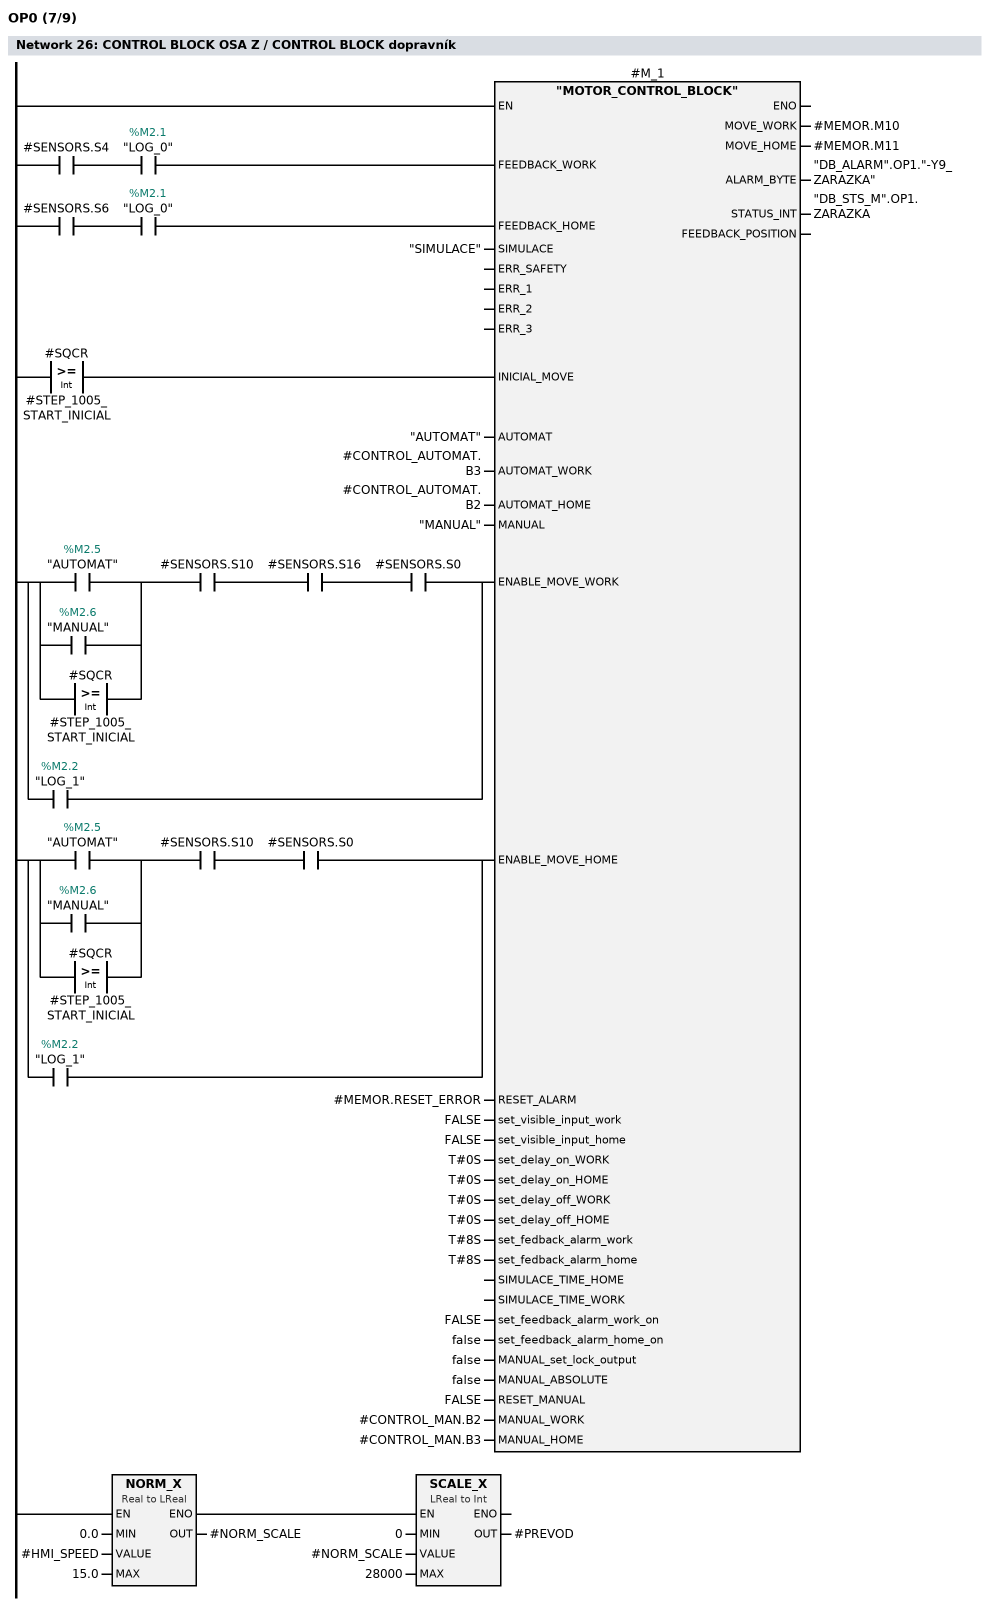
   RUNG wire#powerrail
      #M_1(FEEDBACK_WORK := wire#w1, FEEDBACK_HOME := wire#w2, INICIAL_MOVE := wire#w3, ENABLE_MOVE_WORK := wire#w5, ENABLE_MOVE_HOME := wire#w7, SIMULACE := "SIMULACE", ERR_SAFETY :=, ERR_1 :=, ERR_2 :=, ERR_3 :=, AUTOMAT := "AUTOMAT", AUTOMAT_WORK := #CONTROL_AUTOMAT.B3, AUTOMAT_HOME := #CONTROL_AUTOMAT.B2, MANUAL := "MANUAL", RESET_ALARM := #MEMOR.RESET_ERROR, set_visible_input_work := FALSE, set_visible_input_home := FALSE, set_delay_on_WORK := T#0S, set_delay_on_HOME := T#0S, set_delay_off_WORK := T#0S, set_delay_off_HOME := T#0S, set_fedback_alarm_work := T#8S, set_fedback_alarm_home := T#8S, SIMULACE_TIME_HOME :=, SIMULACE_TIME_WORK :=, set_feedback_alarm_work_on := FALSE, set_feedback_alarm_home_on := false, MANUAL_set_lock_output := false, MANUAL_ABSOLUTE := false, RESET_MANUAL := FALSE, MANUAL_WORK := #CONTROL_MAN.B2, MANUAL_HOME := #CONTROL_MAN.B3, MOVE_WORK => #MEMOR.M10, MOVE_HOME => #MEMOR.M11, ALARM_BYTE => "DB_ALARM".OP1."-Y9_ZARAZKA", STATUS_INT => "DB_STS_M".OP1.ZARAZKA, FEEDBACK_POSITION =>)
   END_RUNG
   RUNG wire#powerrail
      Contact( #SENSORS.S4 )
      Contact( "LOG_0" )
   END_RUNG wire#w1
   RUNG wire#powerrail
      Contact( #SENSORS.S6 )
      Contact( "LOG_0" )
   END_RUNG wire#w2
   RUNG wire#powerrail
      { S7_Templates := "SrcType := Int" } GE_Contact(in1 := #SQCR, in2 := #STEP_1005_START_INICIAL)
   END_RUNG wire#w3
   RUNG wire#powerrail
      Contact( "AUTOMAT" )
      wire#w4
      Contact( #SENSORS.S10 )
      Contact( #SENSORS.S16 )
      Contact( #SENSORS.S0 )
   END_RUNG wire#w5
   RUNG wire#powerrail
      Contact( "MANUAL" )
   END_RUNG wire#w4
   RUNG wire#powerrail
      { S7_Templates := "SrcType := Int" } GE_Contact(in1 := #SQCR, in2 := #STEP_1005_START_INICIAL)
   END_RUNG wire#w4
   RUNG wire#powerrail
      Contact( "LOG_1" )
   END_RUNG wire#w5
   RUNG wire#powerrail
      Contact( "AUTOMAT" )
      wire#w6
      Contact( #SENSORS.S10 )
      Contact( #SENSORS.S0 )
   END_RUNG wire#w7
   RUNG wire#powerrail
      Contact( "MANUAL" )
   END_RUNG wire#w6
   RUNG wire#powerrail
      { S7_Templates := "SrcType := Int" } GE_Contact(in1 := #SQCR, in2 := #STEP_1005_START_INICIAL)
   END_RUNG wire#w6
   RUNG wire#powerrail
      Contact( "LOG_1" )
   END_RUNG wire#w7
   RUNG wire#powerrail
      { S7_Templates := "[SrcType := Real, DestType := LReal]" } Normalize(min := 0.0, value := #HMI_SPEED, max := 15.0, out => #NORM_SCALE)
      { S7_Templates := "[SrcType := LReal, DestType := Int]" } Scale(min := 0, value := #NORM_SCALE, max := 28000, out => #PREVOD)
   END_RUNG
   // the same network as SCL:
   #M_1(FEEDBACK_WORK := #SENSORS.S4 AND "LOG_0",   // "MOTOR_CONTROL_BLOCK"
        FEEDBACK_HOME := #SENSORS.S6 AND "LOG_0",
        SIMULACE := "SIMULACE",
        INICIAL_MOVE := #SQCR >= #STEP_1005_START_INICIAL,
        AUTOMAT := "AUTOMAT",
        AUTOMAT_WORK := #CONTROL_AUTOMAT.B3,
        AUTOMAT_HOME := #CONTROL_AUTOMAT.B2,
        MANUAL := "MANUAL",
        ENABLE_MOVE_WORK := (("AUTOMAT" OR "MANUAL" OR (#SQCR >= #STEP_1005_START_INICIAL)) AND #SENSORS.S10 AND #SENSORS.S16 AND #SENSORS.S0) OR "LOG_1",
        ENABLE_MOVE_HOME := (("AUTOMAT" OR "MANUAL" OR (#SQCR >= #STEP_1005_START_INICIAL)) AND #SENSORS.S10 AND #SENSORS.S0) OR "LOG_1",
        RESET_ALARM := #MEMOR.RESET_ERROR,
        set_visible_input_work := FALSE,
        set_visible_input_home := FALSE,
        set_delay_on_WORK := T#0S,
        set_delay_on_HOME := T#0S,
        set_delay_off_WORK := T#0S,
        set_delay_off_HOME := T#0S,
        set_fedback_alarm_work := T#8S,
        set_fedback_alarm_home := T#8S,
        set_feedback_alarm_work_on := FALSE,
        set_feedback_alarm_home_on := false,
        MANUAL_set_lock_output := false,
        MANUAL_ABSOLUTE := false,
        RESET_MANUAL := FALSE,
        MANUAL_WORK := #CONTROL_MAN.B2,
        MANUAL_HOME := #CONTROL_MAN.B3,
        MOVE_WORK => #MEMOR.M10,
        MOVE_HOME => #MEMOR.M11,
        ALARM_BYTE => "DB_ALARM".OP1."-Y9_ZARAZKA",
        STATUS_INT => "DB_STS_M".OP1.ZARAZKA);
   #NORM_SCALE := NORM_X(MIN := 0.0, VALUE := #HMI_SPEED, MAX := 15.0);
   #PREVOD := SCALE_X(MIN := 0, VALUE := #NORM_SCALE, MAX := 28000);
END_REGION

REGION Network 27: CONTROL BLOCK ARETACE HLAVY / CONTROL BLOCK dveře laser
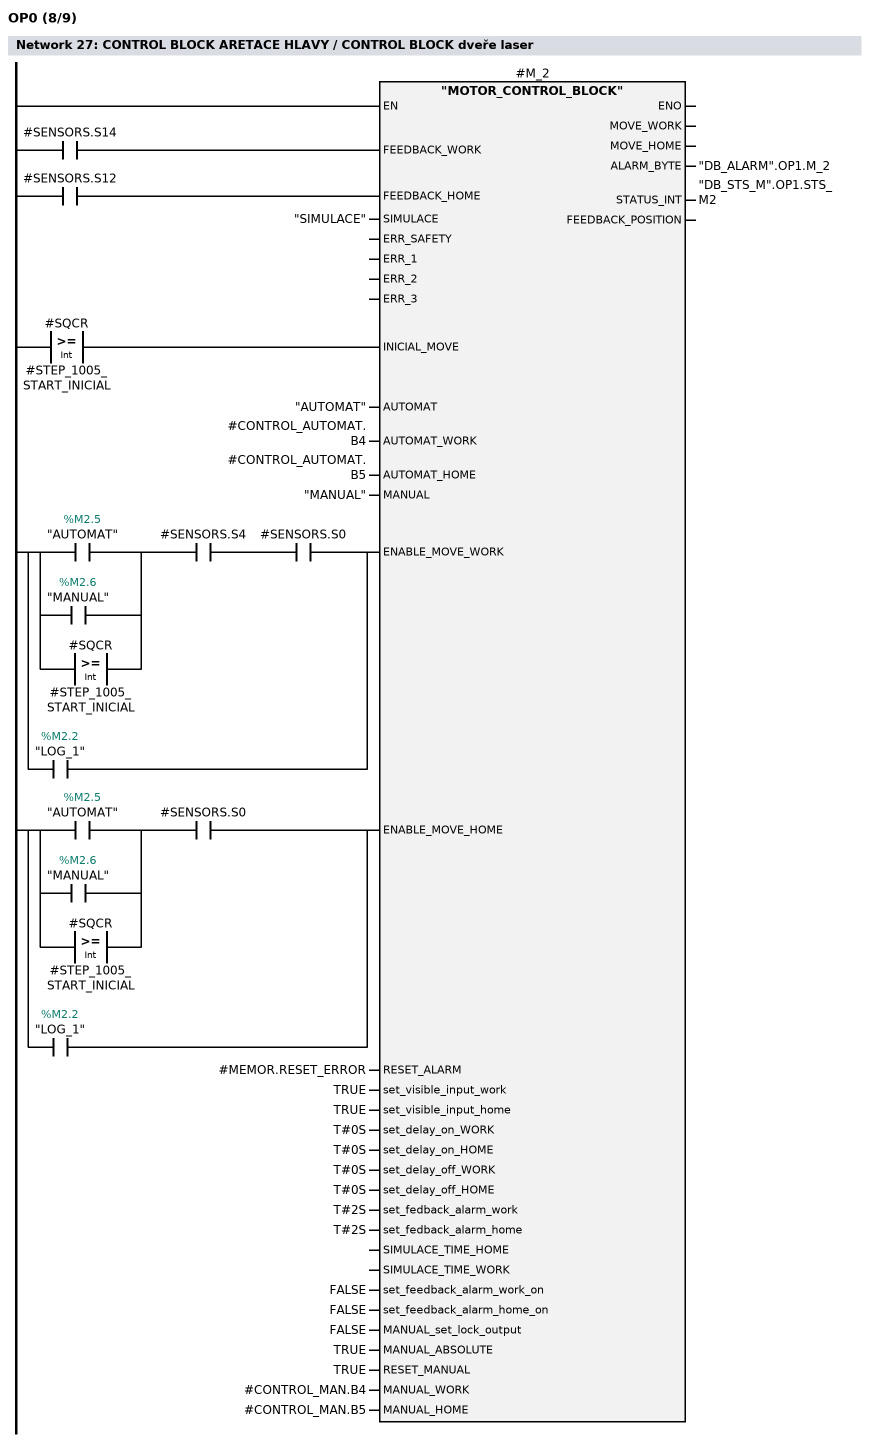
   RUNG wire#powerrail
      #M_2(FEEDBACK_WORK := wire#w1, FEEDBACK_HOME := wire#w2, INICIAL_MOVE := wire#w3, ENABLE_MOVE_WORK := wire#w5, ENABLE_MOVE_HOME := wire#w7, SIMULACE := "SIMULACE", ERR_SAFETY :=, ERR_1 :=, ERR_2 :=, ERR_3 :=, AUTOMAT := "AUTOMAT", AUTOMAT_WORK := #CONTROL_AUTOMAT.B4, AUTOMAT_HOME := #CONTROL_AUTOMAT.B5, MANUAL := "MANUAL", RESET_ALARM := #MEMOR.RESET_ERROR, set_visible_input_work := TRUE, set_visible_input_home := TRUE, set_delay_on_WORK := T#0S, set_delay_on_HOME := T#0S, set_delay_off_WORK := T#0S, set_delay_off_HOME := T#0S, set_fedback_alarm_work := T#2S, set_fedback_alarm_home := T#2S, SIMULACE_TIME_HOME :=, SIMULACE_TIME_WORK :=, set_feedback_alarm_work_on := FALSE, set_feedback_alarm_home_on := FALSE, MANUAL_set_lock_output := FALSE, MANUAL_ABSOLUTE := TRUE, RESET_MANUAL := TRUE, MANUAL_WORK := #CONTROL_MAN.B4, MANUAL_HOME := #CONTROL_MAN.B5, MOVE_WORK =>, MOVE_HOME =>, ALARM_BYTE => "DB_ALARM".OP1.M_2, STATUS_INT => "DB_STS_M".OP1.STS_M2, FEEDBACK_POSITION =>)
   END_RUNG
   RUNG wire#powerrail
      Contact( #SENSORS.S14 )
   END_RUNG wire#w1
   RUNG wire#powerrail
      Contact( #SENSORS.S12 )
   END_RUNG wire#w2
   RUNG wire#powerrail
      { S7_Templates := "SrcType := Int" } GE_Contact(in1 := #SQCR, in2 := #STEP_1005_START_INICIAL)
   END_RUNG wire#w3
   RUNG wire#powerrail
      Contact( "AUTOMAT" )
      wire#w4
      Contact( #SENSORS.S4 )
      Contact( #SENSORS.S0 )
   END_RUNG wire#w5
   RUNG wire#powerrail
      Contact( "MANUAL" )
   END_RUNG wire#w4
   RUNG wire#powerrail
      { S7_Templates := "SrcType := Int" } GE_Contact(in1 := #SQCR, in2 := #STEP_1005_START_INICIAL)
   END_RUNG wire#w4
   RUNG wire#powerrail
      Contact( "LOG_1" )
   END_RUNG wire#w5
   RUNG wire#powerrail
      Contact( "AUTOMAT" )
      wire#w6
      Contact( #SENSORS.S0 )
   END_RUNG wire#w7
   RUNG wire#powerrail
      Contact( "MANUAL" )
   END_RUNG wire#w6
   RUNG wire#powerrail
      { S7_Templates := "SrcType := Int" } GE_Contact(in1 := #SQCR, in2 := #STEP_1005_START_INICIAL)
   END_RUNG wire#w6
   RUNG wire#powerrail
      Contact( "LOG_1" )
   END_RUNG wire#w7
   // the same network as SCL:
   #M_2(FEEDBACK_WORK := #SENSORS.S14,   // "MOTOR_CONTROL_BLOCK"
        FEEDBACK_HOME := #SENSORS.S12,
        SIMULACE := "SIMULACE",
        INICIAL_MOVE := #SQCR >= #STEP_1005_START_INICIAL,
        AUTOMAT := "AUTOMAT",
        AUTOMAT_WORK := #CONTROL_AUTOMAT.B4,
        AUTOMAT_HOME := #CONTROL_AUTOMAT.B5,
        MANUAL := "MANUAL",
        ENABLE_MOVE_WORK := (("AUTOMAT" OR "MANUAL" OR (#SQCR >= #STEP_1005_START_INICIAL)) AND #SENSORS.S4 AND #SENSORS.S0) OR "LOG_1",
        ENABLE_MOVE_HOME := (("AUTOMAT" OR "MANUAL" OR (#SQCR >= #STEP_1005_START_INICIAL)) AND #SENSORS.S0) OR "LOG_1",
        RESET_ALARM := #MEMOR.RESET_ERROR,
        set_visible_input_work := TRUE,
        set_visible_input_home := TRUE,
        set_delay_on_WORK := T#0S,
        set_delay_on_HOME := T#0S,
        set_delay_off_WORK := T#0S,
        set_delay_off_HOME := T#0S,
        set_fedback_alarm_work := T#2S,
        set_fedback_alarm_home := T#2S,
        set_feedback_alarm_work_on := FALSE,
        set_feedback_alarm_home_on := FALSE,
        MANUAL_set_lock_output := FALSE,
        MANUAL_ABSOLUTE := TRUE,
        RESET_MANUAL := TRUE,
        MANUAL_WORK := #CONTROL_MAN.B4,
        MANUAL_HOME := #CONTROL_MAN.B5,
        ALARM_BYTE => "DB_ALARM".OP1.M_2,
        STATUS_INT => "DB_STS_M".OP1.STS_M2);
END_REGION

REGION Network 28: EXTERNAL_TRIGER
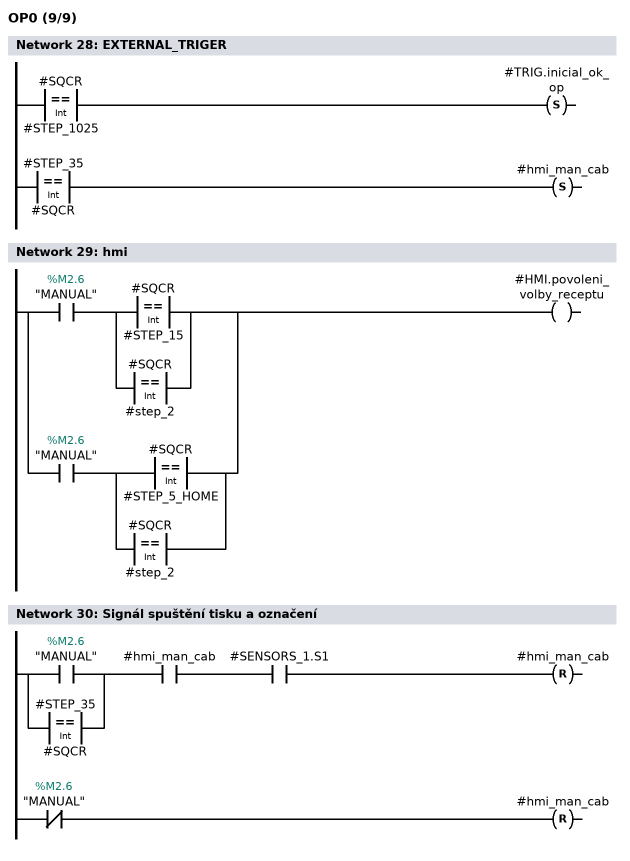
   RUNG wire#powerrail
      { S7_Templates := "SrcType := Int" } EQ_Contact(in1 := #SQCR, in2 := #STEP_1025)
      S_Coil( #TRIG.inicial_ok_op )
   END_RUNG
   RUNG wire#powerrail
      { S7_Templates := "SrcType := Int" } EQ_Contact(in1 := #STEP_35, in2 := #SQCR)
      S_Coil( #hmi_man_cab )
   END_RUNG
   // the same network as SCL:
   IF #SQCR = #STEP_1025 THEN #TRIG.inicial_ok_op := TRUE; END_IF;
   IF #STEP_35 = #SQCR THEN #hmi_man_cab := TRUE; END_IF;
END_REGION

REGION Network 29: hmi
   RUNG wire#powerrail
      Contact( "MANUAL" )
      wire#w1
      { S7_Templates := "SrcType := Int" } EQ_Contact(in1 := #SQCR, in2 := #STEP_15)
      wire#w2
      Coil( #HMI.povoleni_volby_receptu )
   END_RUNG
   RUNG wire#w1
      { S7_Templates := "SrcType := Int" } EQ_Contact(in1 := #SQCR, in2 := #step_2)
   END_RUNG wire#w2
   RUNG wire#powerrail
      Contact( "MANUAL" )
      wire#w3
      { S7_Templates := "SrcType := Int" } EQ_Contact(in1 := #SQCR, in2 := #STEP_5_HOME)
   END_RUNG wire#w2
   RUNG wire#w3
      { S7_Templates := "SrcType := Int" } EQ_Contact(in1 := #SQCR, in2 := #step_2)
   END_RUNG wire#w2
   // the same network as SCL:
   #HMI.povoleni_volby_receptu := ("MANUAL" AND ((#SQCR = #STEP_15) OR (#SQCR = #step_2))) OR ("MANUAL" AND ((#SQCR = #STEP_5_HOME) OR (#SQCR = #step_2)));
END_REGION

REGION Network 30: Signál spuštění tisku a označení
   RUNG wire#powerrail
      Contact( "MANUAL" )
      wire#w1
      Contact( #hmi_man_cab )
      Contact( #SENSORS_1.S1 )
      R_Coil( #hmi_man_cab )
   END_RUNG
   RUNG wire#powerrail
      { S7_Templates := "SrcType := Int" } EQ_Contact(in1 := #STEP_35, in2 := #SQCR)
   END_RUNG wire#w1
   RUNG wire#powerrail
      I_Contact( "MANUAL" )
      R_Coil( #hmi_man_cab )
   END_RUNG
   // the same network as SCL:
   IF ("MANUAL" OR (#STEP_35 = #SQCR)) AND #hmi_man_cab AND #SENSORS_1.S1 THEN #hmi_man_cab := FALSE; END_IF;
   IF NOT "MANUAL" THEN #hmi_man_cab := FALSE; END_IF;
END_REGION
END_FUNCTION_BLOCK

FUNCTION_BLOCK "OVLADANI_LASER"   // FB400, LAD
{ S7_Optimized_Access := 'TRUE' }
// stored: AutoNumber false, MemoryReserve 100, SetENOAutomatically false
   VAR
      SQCR : Int;
      SQCR_WHILE : Int;
      SET_WHILE : Bool;
      NAZEV_PROGRAMU : String[20];
      DELKA_STRINGU : Int;
      CHAR_K_ZAPISU : Array[0..71] of Char;
   END_VAR
   VAR CONSTANT
      STEP_0 : Int := 0;
      STEP_5 : Int := 5;
      STEP_10 : Int := 10;
      STEP_15 : Int := 15;
      STEP_20 : Int := 20;
      STEP_25 : Int := 25;
      STEP_30 : Int := 30;
      STEP_35 : Int := 35;
      STEP_40 : Int := 40;
      STEP_45 : Int := 45;
      STEP_50 : Int := 50;
      STEP_55 : Int := 55;
      STEP_60 : Int := 60;
      STEP_65 : Int := 65;
      STEP_70 : Int := 70;
      STEP_75 : Int := 75;
      STEP_80 : Int := 80;
      STEP_85 : Int := 85;
      STEP_90 : Int := 90;
      STEP_95 : Int := 95;
      STEP_100 : Int := 100;
   END_VAR
BEGIN

REGION Network 1
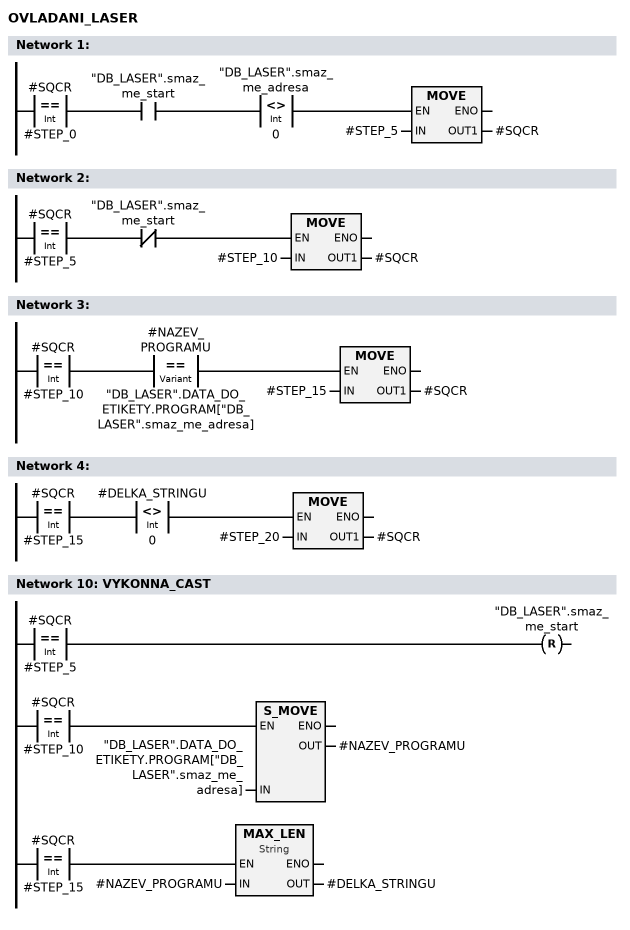
   RUNG wire#powerrail
      { S7_Templates := "SrcType := Int" } EQ_Contact(in1 := #SQCR, in2 := #STEP_0)
      Contact( "DB_LASER".smaz_me_start )
      { S7_Templates := "SrcType := Int" } NE_Contact(in1 := "DB_LASER".smaz_me_adresa, in2 := 0)
      Move(in := #STEP_5, out1 => #SQCR)
   END_RUNG
   // the same network as SCL:
   IF (#SQCR = #STEP_0) AND "DB_LASER".smaz_me_start AND ("DB_LASER".smaz_me_adresa <> 0) THEN
       #SQCR := #STEP_5;
   END_IF;
END_REGION

REGION Network 2
   RUNG wire#powerrail
      { S7_Templates := "SrcType := Int" } EQ_Contact(in1 := #SQCR, in2 := #STEP_5)
      I_Contact( "DB_LASER".smaz_me_start )
      Move(in := #STEP_10, out1 => #SQCR)
   END_RUNG
   // the same network as SCL:
   IF (#SQCR = #STEP_5) AND NOT "DB_LASER".smaz_me_start THEN #SQCR := #STEP_10; END_IF;
END_REGION

REGION Network 3
   RUNG wire#powerrail
      { S7_Templates := "SrcType := Int" } EQ_Contact(in1 := #SQCR, in2 := #STEP_10)
      { S7_Templates := "SrcType := Variant" } EQ_Contact(in1 := #NAZEV_PROGRAMU, in2 := "DB_LASER".DATA_DO_ETIKETY.PROGRAM["DB_LASER".smaz_me_adresa])
      Move(in := #STEP_15, out1 => #SQCR)
   END_RUNG
   // the same network as SCL:
   IF (#SQCR = #STEP_10) AND (#NAZEV_PROGRAMU = "DB_LASER".DATA_DO_ETIKETY.PROGRAM["DB_LASER".smaz_me_adresa]) THEN
       #SQCR := #STEP_15;
   END_IF;
END_REGION

REGION Network 4
   RUNG wire#powerrail
      { S7_Templates := "SrcType := Int" } EQ_Contact(in1 := #SQCR, in2 := #STEP_15)
      { S7_Templates := "SrcType := Int" } NE_Contact(in1 := #DELKA_STRINGU, in2 := 0)
      Move(in := #STEP_20, out1 => #SQCR)
   END_RUNG
   // the same network as SCL:
   IF (#SQCR = #STEP_15) AND (#DELKA_STRINGU <> 0) THEN #SQCR := #STEP_20; END_IF;
END_REGION

REGION Network 5: STEP_20 SCL NETVORK X
END_REGION

REGION Network 10: VYKONNA_CAST
   IF #SQCR = #STEP_5 THEN "DB_LASER".smaz_me_start := FALSE; END_IF;
   IF #SQCR = #STEP_10 THEN
       #NAZEV_PROGRAMU := "DB_LASER".DATA_DO_ETIKETY.PROGRAM["DB_LASER".smaz_me_adresa];
   END_IF;
   IF #SQCR = #STEP_15 THEN MAX_LEN(in := #NAZEV_PROGRAMU, out => #DELKA_STRINGU); END_IF;
END_REGION

REGION Network 12 (SCL)
   IF #SQCR = #STEP_20 THEN
       // zapsani počátečního znaku 
       #CHAR_K_ZAPISU[0] := "DB_LASER".DATA_DO_DAT.ZAVORKA_P;



       // vytvoření prdelky k názvu programu z laseru
       #CHAR_K_ZAPISU[#DELKA_STRINGU + 1] := "DB_LASER".DATA_DO_DAT.XLP[0];
       #CHAR_K_ZAPISU[#DELKA_STRINGU + 2] := "DB_LASER".DATA_DO_DAT.XLP[1];
       #CHAR_K_ZAPISU[#DELKA_STRINGU + 3] := "DB_LASER".DATA_DO_DAT.XLP[2];
       #CHAR_K_ZAPISU[#DELKA_STRINGU + 4] := "DB_LASER".DATA_DO_DAT.XLP[3];
       #CHAR_K_ZAPISU[#DELKA_STRINGU + 5] := "DB_LASER".DATA_DO_DAT.ZAVORKA_P;

       // dinamický zápis názvu podle délky stringu 
       WHILE #SET_WHILE DO
           IF #SQCR_WHILE > #DELKA_STRINGU THEN
               #SQCR_WHILE := 0;
               #SET_WHILE := FALSE;
               #SQCR := #STEP_25;
           ELSE
               #SQCR_WHILE := #SQCR_WHILE + 1;
           END_IF;
           #CHAR_K_ZAPISU[#SQCR_WHILE + 1] := #NAZEV_PROGRAMU[#SQCR_WHILE];
       END_WHILE;

   END_IF;
END_REGION
END_FUNCTION_BLOCK

FUNCTION "FC_PocetChyb" : Int
{ S7_Optimized_Access := 'TRUE' }
VERSION : 0.1
   VAR_INPUT 
      A : String;
      B : String;
   END_VAR

   VAR_TEMP 
      la : Int;
      lb : Int;
      i : Int;
      j : Int;
      v : Int;
      prev : Array[0..40] of Int;
      cur : Array[0..40] of Int;
   END_VAR


BEGIN
	// Pocet chyb mezi texty A a B (kolik znaku zamenit / vlozit / smazat).
	// 0 = texty jsou shodne. Porovnava se max. 40 znaku kvuli dobe cyklu.
	#la := MIN(IN1 := LEN(#A), IN2 := 40);
	#lb := MIN(IN1 := LEN(#B), IN2 := 40);
	
	FOR #j := 0 TO #lb DO
	    #prev[#j] := #j;
	END_FOR;
	
	FOR #i := 1 TO #la DO
	    #cur[0] := #i;
	    FOR #j := 1 TO #lb DO
	        #v := #prev[#j - 1];                // shoda / zamena znaku
	        IF #A[#i] <> #B[#j] THEN
	            #v := #v + 1;
	        END_IF;
	        IF #prev[#j] + 1 < #v THEN          // znak navic
	            #v := #prev[#j] + 1;
	        END_IF;
	        IF #cur[#j - 1] + 1 < #v THEN       // chybejici znak
	            #v := #cur[#j - 1] + 1;
	        END_IF;
	        #cur[#j] := #v;
	    END_FOR;
	    FOR #j := 0 TO #lb DO
	        #prev[#j] := #cur[#j];
	    END_FOR;
	END_FOR;
	
	#FC_PocetChyb := #prev[#lb];
END_FUNCTION

DATA_BLOCK "OP1_DB"   // DB50
// stored: AutoNumber false, InstanceOfName OP1, InstanceOfType FB
"OP1"
BEGIN
END_DATA_BLOCK

DATA_BLOCK "OP2_DB"   // DB1
// stored: InstanceOfName OP2, InstanceOfType FB
"OP2"
BEGIN
END_DATA_BLOCK

DATA_BLOCK "iDB_CamManual"   // DB9
// stored: InstanceOfName FB_CamManual, InstanceOfType FB
"FB_CamManual"
BEGIN
END_DATA_BLOCK

DATA_BLOCK "CONTROL_LINE_DB"   // DB27
// stored: AutoNumber false, InstanceOfName CONTROL_LINE, InstanceOfType FB
"CONTROL_LINE"
BEGIN
END_DATA_BLOCK

DATA_BLOCK "OVLADANI_LASER_DB"   // DB400
// stored: AutoNumber false, InstanceOfName OVLADANI_LASER, InstanceOfType FB
"OVLADANI_LASER"
BEGIN
END_DATA_BLOCK
